Fanuc KAREL source: kc00002.KL

-- PROVISIONAL review KL for V1013-1; original PC SHA256 6b39b8591156d7d7cd8d995d1a04dcfe2f6d2b66c2ae0d3e75acbdd42b76922f
-- Incomplete behavior may be omitted. Consult companion uncertainty JSON. Do not deploy.
PROGRAM KC00002
%NOLOCKGROUP
BEGIN
  -- UNRESOLVED_PC offsets 5-33; opcodes 27,22,22,22,22,31
  -- UNRESOLVED_PC offsets 38-42; opcodes 7F
END KC00002
